(* IEC 61131-3 sources: horner-cscape-mcp/artifacts/projects/Fail_Undeclared_Location_Proj/pous, 1 file *)

(* ---- POU_UndeclaredVar.st ---- *)
PROGRAM POU_UndeclaredVar
VAR
    ValidCounter : INT := 0;
END_VAR

PhantomOutput := 99;
END_PROGRAM
